screen "D_Bar_1" 1280x800
   Bar "Static" at 6,4 size 40x120
   TextField "Label_Static" at 6,156 size 55x22; Text 'Static'
   Bar "A_Range" at 98,4 size 40x120
      Appearance <- "D_Range"
   TextField "Label_A_Range" at 98,156 size 79x22; Text 'A_Range'
   Bar "A_Flash" at 190,4 size 40x120
      Appearance <- "D_Range"
   TextField "Label_A_Flash" at 190,156 size 72x22; Text 'A_Flash'
   Bar "A_Bit" at 282,4 size 40x120
      Appearance <- "D_Bool"
   TextField "Label_A_Bit" at 282,156 size 51x22; Text 'A_Bit'
   Bar "A_Bits" at 374,4 size 40x120
      Appearance <- "D_Bits"
   TextField "Label_A_Bits" at 374,156 size 60x22; Text 'A_Bits'
   Bar "V_Range" at 466,4 size 40x120
      Visibility <- "D_Range"
   TextField "Label_V_Range" at 466,156 size 79x22; Text 'V_Range'
   Bar "V_Bit" at 558,4 size 40x120
      Visibility <- "D_Vis"
   TextField "Label_V_Bit" at 558,156 size 51x22; Text 'V_Bit'
   Bar "M_H" at 650,4 size 40x120
      HorizontalMovement <- "D_Pct"
   TextField "Label_M_H" at 650,156 size 42x22; Text 'M_H'
   Bar "M_V" at 742,4 size 40x120
      VerticalMovement <- "D_Pct"
   TextField "Label_M_V" at 742,156 size 41x22; Text 'M_V'
   Bar "M_D" at 834,4 size 40x120
      DiagonalMovement <- "D_Pct"
   TextField "Label_M_D" at 834,156 size 42x22; Text 'M_D'
   Bar "M_Direct" at 926,4 size 40x120
      DirectMovement <- "D_X"
      DirectMovement <- "D_Y"
   TextField "Label_M_Direct" at 926,156 size 82x22; Text 'M_Direct'
   Bar "E_Range" at 1018,4 size 40x120
      ObjectEnable <- "D_Range"
   TextField "Label_E_Range" at 1018,156 size 78x22; Text 'E_Range'
   Bar "E_Bit" at 1110,4 size 40x120
      ObjectEnable <- "D_En"
   TextField "Label_E_Bit" at 1110,156 size 50x22; Text 'E_Bit'
   Bar "PV_Pct" at 6,176 size 40x120
      ProcessValue <- "D_Pct"
   TextField "Label_PV_Pct" at 6,328 size 65x22; Text 'PV_Pct'
   Bar "PV_Real" at 98,176 size 40x120
      ProcessValue <- "D_Real"
   TextField "Label_PV_Real" at 98,328 size 76x22; Text 'PV_Real'
   Bar "PV_BarR" at 190,176 size 40x120
      ProcessValue <- "D_BarR"
   TextField "Label_PV_BarR" at 190,328 size 79x22; Text 'PV_BarR'
   Bar "PV_Pct_0_100" at 282,176 size 40x120; MinimumValue 0; MaximumValue 100
      ProcessValue <- "D_Pct"
   TextField "Label_PV_Pct_0_100" at 282,328 size 131x22; Text 'PV_Pct_0_100'
   Bar "PV_Pct_MaxMin" at 374,176 size 40x120
      ProcessValue <- "D_Pct"
      MaximumValue <- "D_Max"
      MinimumValue <- "D_Min"
   TextField "Label_PV_Pct_MaxMin" at 374,328 size 140x22; Text 'PV_Pct_MaxMin'
   IOField "State" at 4,774 size 60x22; FormatPattern 9
      ProcessValue <- "D_State"
   Button "S1" at 70,774 size 40x22; TextOff 'S1'
      on Click: "SetS1"()
   Button "S2" at 114,774 size 40x22; TextOff 'S2'
      on Click: "SetS2"()
   Button "S3" at 158,774 size 40x22; TextOff 'S3'
      on Click: "SetS3"()
   Button "S4" at 202,774 size 40x22; TextOff 'S4'
      on Click: "SetS4"()
   Button "Next" at 1236,774 size 40x22; TextOff 'Next'
      on Click: ActivateScreen("D_Switch_1", 0)

screen "D_Button_1" 1280x800
   Button "Static" at 6,4 size 100x40; TextOff 'Text'
   TextField "Label_Static" at 6,76 size 55x22; Text 'Static'
   Button "A_Range" at 158,4 size 100x40; TextOff 'Text'
      Appearance <- "D_Range"
   TextField "Label_A_Range" at 158,76 size 79x22; Text 'A_Range'
   Button "A_Flash" at 310,4 size 100x40; TextOff 'Text'
      Appearance <- "D_Range"
   TextField "Label_A_Flash" at 310,76 size 72x22; Text 'A_Flash'
   Button "A_Bit" at 462,4 size 100x40; TextOff 'Text'
      Appearance <- "D_Bool"
   TextField "Label_A_Bit" at 462,76 size 51x22; Text 'A_Bit'
   Button "A_Bits" at 614,4 size 100x40; TextOff 'Text'
      Appearance <- "D_Bits"
   TextField "Label_A_Bits" at 614,76 size 60x22; Text 'A_Bits'
   Button "V_Range" at 766,4 size 100x40; TextOff 'Text'
      Visibility <- "D_Range"
   TextField "Label_V_Range" at 766,76 size 79x22; Text 'V_Range'
   Button "V_Bit" at 918,4 size 100x40; TextOff 'Text'
      Visibility <- "D_Vis"
   TextField "Label_V_Bit" at 918,76 size 51x22; Text 'V_Bit'
   Button "M_H" at 1070,4 size 100x40; TextOff 'Text'
      HorizontalMovement <- "D_Pct"
   TextField "Label_M_H" at 1070,76 size 42x22; Text 'M_H'
   Button "M_V" at 6,96 size 100x40; TextOff 'Text'
      VerticalMovement <- "D_Pct"
   TextField "Label_M_V" at 6,168 size 41x22; Text 'M_V'
   Button "M_D" at 158,96 size 100x40; TextOff 'Text'
      DiagonalMovement <- "D_Pct"
   TextField "Label_M_D" at 158,168 size 42x22; Text 'M_D'
   Button "M_Direct" at 310,96 size 100x40; TextOff 'Text'
      DirectMovement <- "D_X"
      DirectMovement <- "D_Y"
   TextField "Label_M_Direct" at 310,168 size 82x22; Text 'M_Direct'
   Button "E_Range" at 462,96 size 100x40; TextOff 'Text'
      ObjectEnable <- "D_Range"
   TextField "Label_E_Range" at 462,168 size 78x22; Text 'E_Range'
   Button "E_Bit" at 614,96 size 100x40; TextOff 'Text'
      ObjectEnable <- "D_En"
   TextField "Label_E_Bit" at 614,168 size 50x22; Text 'E_Bit'
   IOField "State" at 4,774 size 60x22; FormatPattern 9
      ProcessValue <- "D_State"
   Button "S1" at 70,774 size 40x22; TextOff 'S1'
      on Click: "SetS1"()
   Button "S2" at 114,774 size 40x22; TextOff 'S2'
      on Click: "SetS2"()
   Button "S3" at 158,774 size 40x22; TextOff 'S3'
      on Click: "SetS3"()
   Button "S4" at 202,774 size 40x22; TextOff 'S4'
      on Click: "SetS4"()
   Button "Next" at 1236,774 size 40x22; TextOff 'Next'
      on Click: ActivateScreen("D_SymbolicIOField_1", 0)

screen "D_Circle_1" 1280x800
   TextField "Label_Static" at 6,86 size 55x22; Text 'Static'
   Circle "A_Range" at 108,4 size 50x50
      Appearance <- "D_Range"
   TextField "Label_A_Range" at 108,86 size 79x22; Text 'A_Range'
   Circle "A_Flash" at 210,4 size 50x50
      Appearance <- "D_Range"
   TextField "Label_A_Flash" at 210,86 size 72x22; Text 'A_Flash'
   Circle "A_Bit" at 312,4 size 50x50
      Appearance <- "D_Bool"
   TextField "Label_A_Bit" at 312,86 size 51x22; Text 'A_Bit'
   Circle "A_Bits" at 414,4 size 50x50
      Appearance <- "D_Bits"
   TextField "Label_A_Bits" at 414,86 size 60x22; Text 'A_Bits'
   Circle "V_Range" at 516,4 size 50x50
      Visibility <- "D_Range"
   TextField "Label_V_Range" at 516,86 size 79x22; Text 'V_Range'
   Circle "V_Bit" at 618,4 size 50x50
      Visibility <- "D_Vis"
   TextField "Label_V_Bit" at 618,86 size 51x22; Text 'V_Bit'
   Circle "M_H" at 720,4 size 50x50
      HorizontalMovement <- "D_Pct"
   TextField "Label_M_H" at 720,86 size 42x22; Text 'M_H'
   Circle "M_V" at 822,4 size 50x50
      VerticalMovement <- "D_Pct"
   TextField "Label_M_V" at 822,86 size 41x22; Text 'M_V'
   Circle "M_D" at 924,4 size 50x50
      DiagonalMovement <- "D_Pct"
   TextField "Label_M_D" at 924,86 size 42x22; Text 'M_D'
   Circle "M_Direct" at 1026,4 size 50x50
      DirectMovement <- "D_X"
      DirectMovement <- "D_Y"
   TextField "Label_M_Direct" at 1026,86 size 82x22; Text 'M_Direct'
   Circle "E_Range" at 1128,4 size 50x50
      ObjectEnable <- "D_Range"
   TextField "Label_E_Range" at 1128,86 size 78x22; Text 'E_Range'
   Circle "E_Bit" at 6,106 size 50x50
      ObjectEnable <- "D_En"
   TextField "Label_E_Bit" at 6,188 size 50x22; Text 'E_Bit'
   IOField "State" at 4,774 size 60x22; FormatPattern 9
      ProcessValue <- "D_State"
   Button "S1" at 70,774 size 40x22; TextOff 'S1'
      on Click: "SetS1"()
   Button "S2" at 114,774 size 40x22; TextOff 'S2'
      on Click: "SetS2"()
   Button "S3" at 158,774 size 40x22; TextOff 'S3'
      on Click: "SetS3"()
   Button "S4" at 202,774 size 40x22; TextOff 'S4'
      on Click: "SetS4"()
   Button "Next" at 1236,774 size 40x22; TextOff 'Next'
      on Click: ActivateScreen("D_Rectangle_1", 0)

screen "D_Clock_1" 1280x800
   Clock "Static" at 6,4 size 150x150
   TextField "Label_Static" at 6,186 size 55x22; Text 'Static'
   Clock "A_Range" at 208,4 size 150x150
      Appearance <- "D_Range"
   TextField "Label_A_Range" at 208,186 size 79x22; Text 'A_Range'
   Clock "A_Flash" at 410,4 size 150x150
      Appearance <- "D_Range"
   TextField "Label_A_Flash" at 410,186 size 72x22; Text 'A_Flash'
   Clock "A_Bit" at 612,4 size 150x150
      Appearance <- "D_Bool"
   TextField "Label_A_Bit" at 612,186 size 51x22; Text 'A_Bit'
   Clock "A_Bits" at 814,4 size 150x150
      Appearance <- "D_Bits"
   TextField "Label_A_Bits" at 814,186 size 60x22; Text 'A_Bits'
   Clock "V_Range" at 1016,4 size 150x150
      Visibility <- "D_Range"
   TextField "Label_V_Range" at 1016,186 size 79x22; Text 'V_Range'
   Clock "V_Bit" at 6,206 size 150x150
      Visibility <- "D_Vis"
   TextField "Label_V_Bit" at 6,388 size 51x22; Text 'V_Bit'
   Clock "M_H" at 208,206 size 150x150
      HorizontalMovement <- "D_Pct"
   TextField "Label_M_H" at 208,388 size 42x22; Text 'M_H'
   Clock "M_V" at 410,206 size 150x150
      VerticalMovement <- "D_Pct"
   TextField "Label_M_V" at 410,388 size 41x22; Text 'M_V'
   Clock "M_D" at 612,206 size 150x150
      DiagonalMovement <- "D_Pct"
   TextField "Label_M_D" at 612,388 size 42x22; Text 'M_D'
   Clock "M_Direct" at 814,206 size 150x150
      DirectMovement <- "D_X"
      DirectMovement <- "D_Y"
   TextField "Label_M_Direct" at 814,388 size 82x22; Text 'M_Direct'
   Clock "E_Range" at 1016,206 size 150x150
      ObjectEnable <- "D_Range"
   TextField "Label_E_Range" at 1016,388 size 78x22; Text 'E_Range'
   Clock "E_Bit" at 6,408 size 150x150
      ObjectEnable <- "D_En"
   TextField "Label_E_Bit" at 6,590 size 50x22; Text 'E_Bit'
   IOField "State" at 4,774 size 60x22; FormatPattern 9
      ProcessValue <- "D_State"
   Button "S1" at 70,774 size 40x22; TextOff 'S1'
      on Click: "SetS1"()
   Button "S2" at 114,774 size 40x22; TextOff 'S2'
      on Click: "SetS2"()
   Button "S3" at 158,774 size 40x22; TextOff 'S3'
      on Click: "SetS3"()
   Button "S4" at 202,774 size 40x22; TextOff 'S4'
      on Click: "SetS4"()
   Button "Next" at 1236,774 size 40x22; TextOff 'Next'
      on Click: ActivateScreen("D_Line_1", 0)

screen "D_DateTimeField_1" 1280x800
   DateTimeField "Static" at 6,4 size 189x26
   TextField "Label_Static" at 6,66 size 55x22; Text 'Static'
   DateTimeField "A_Range" at 218,4 size 189x26
      Appearance <- "D_Range"
   TextField "Label_A_Range" at 218,66 size 79x22; Text 'A_Range'
   DateTimeField "A_Flash" at 430,4 size 189x26
      Appearance <- "D_Range"
   TextField "Label_A_Flash" at 430,66 size 72x22; Text 'A_Flash'
   DateTimeField "A_Bit" at 642,4 size 189x26
      Appearance <- "D_Bool"
   TextField "Label_A_Bit" at 642,66 size 51x22; Text 'A_Bit'
   DateTimeField "A_Bits" at 854,4 size 189x26
      Appearance <- "D_Bits"
   TextField "Label_A_Bits" at 854,66 size 60x22; Text 'A_Bits'
   DateTimeField "V_Range" at 1066,4 size 189x26
      Visibility <- "D_Range"
   TextField "Label_V_Range" at 1066,66 size 79x22; Text 'V_Range'
   DateTimeField "V_Bit" at 6,86 size 189x26
      Visibility <- "D_Vis"
   TextField "Label_V_Bit" at 6,148 size 51x22; Text 'V_Bit'
   DateTimeField "M_H" at 218,86 size 189x26
      HorizontalMovement <- "D_Pct"
   TextField "Label_M_H" at 218,148 size 42x22; Text 'M_H'
   DateTimeField "M_V" at 430,86 size 189x26
      VerticalMovement <- "D_Pct"
   TextField "Label_M_V" at 430,148 size 41x22; Text 'M_V'
   DateTimeField "M_D" at 642,86 size 189x26
      DiagonalMovement <- "D_Pct"
   TextField "Label_M_D" at 642,148 size 42x22; Text 'M_D'
   DateTimeField "M_Direct" at 854,86 size 189x26
      DirectMovement <- "D_X"
      DirectMovement <- "D_Y"
   TextField "Label_M_Direct" at 854,148 size 82x22; Text 'M_Direct'
   DateTimeField "E_Range" at 1066,86 size 189x26
      ObjectEnable <- "D_Range"
   TextField "Label_E_Range" at 1066,148 size 78x22; Text 'E_Range'
   DateTimeField "E_Bit" at 6,168 size 189x26
      ObjectEnable <- "D_En"
   TextField "Label_E_Bit" at 6,230 size 50x22; Text 'E_Bit'
   DateTimeField "PV_DateTime" at 218,168 size 189x26
      ProcessValue <- "D_DateTime"
   TextField "Label_PV_DateTime" at 218,230 size 117x22; Text 'PV_DateTime'
   IOField "State" at 4,774 size 60x22; FormatPattern 9
      ProcessValue <- "D_State"
   Button "S1" at 70,774 size 40x22; TextOff 'S1'
      on Click: "SetS1"()
   Button "S2" at 114,774 size 40x22; TextOff 'S2'
      on Click: "SetS2"()
   Button "S3" at 158,774 size 40x22; TextOff 'S3'
      on Click: "SetS3"()
   Button "S4" at 202,774 size 40x22; TextOff 'S4'
      on Click: "SetS4"()
   Button "Next" at 1236,774 size 40x22; TextOff 'Next'
      on Click: ActivateScreen("D_Bar_1", 0)

screen "D_Ellipse_1" 1280x800
   TextField "Label_Static" at 6,86 size 55x22; Text 'Static'
   Ellipse "A_Range" at 158,4 size 100x50
      Appearance <- "D_Range"
   TextField "Label_A_Range" at 158,86 size 79x22; Text 'A_Range'
   Ellipse "A_Flash" at 310,4 size 100x50
      Appearance <- "D_Range"
   TextField "Label_A_Flash" at 310,86 size 72x22; Text 'A_Flash'
   Ellipse "A_Bit" at 462,4 size 100x50
      Appearance <- "D_Bool"
   TextField "Label_A_Bit" at 462,86 size 51x22; Text 'A_Bit'
   Ellipse "A_Bits" at 614,4 size 100x50
      Appearance <- "D_Bits"
   TextField "Label_A_Bits" at 614,86 size 60x22; Text 'A_Bits'
   Ellipse "V_Range" at 766,4 size 100x50
      Visibility <- "D_Range"
   TextField "Label_V_Range" at 766,86 size 79x22; Text 'V_Range'
   Ellipse "V_Bit" at 918,4 size 100x50
      Visibility <- "D_Vis"
   TextField "Label_V_Bit" at 918,86 size 51x22; Text 'V_Bit'
   Ellipse "M_H" at 1070,4 size 100x50
      HorizontalMovement <- "D_Pct"
   TextField "Label_M_H" at 1070,86 size 42x22; Text 'M_H'
   Ellipse "M_V" at 6,106 size 100x50
      VerticalMovement <- "D_Pct"
   TextField "Label_M_V" at 6,188 size 41x22; Text 'M_V'
   Ellipse "M_D" at 158,106 size 100x50
      DiagonalMovement <- "D_Pct"
   TextField "Label_M_D" at 158,188 size 42x22; Text 'M_D'
   Ellipse "M_Direct" at 310,106 size 100x50
      DirectMovement <- "D_X"
      DirectMovement <- "D_Y"
   TextField "Label_M_Direct" at 310,188 size 82x22; Text 'M_Direct'
   Ellipse "E_Range" at 462,106 size 100x50
      ObjectEnable <- "D_Range"
   TextField "Label_E_Range" at 462,188 size 78x22; Text 'E_Range'
   Ellipse "E_Bit" at 614,106 size 100x50
      ObjectEnable <- "D_En"
   TextField "Label_E_Bit" at 614,188 size 50x22; Text 'E_Bit'
   IOField "State" at 4,774 size 60x22; FormatPattern 9
      ProcessValue <- "D_State"
   Button "S1" at 70,774 size 40x22; TextOff 'S1'
      on Click: "SetS1"()
   Button "S2" at 114,774 size 40x22; TextOff 'S2'
      on Click: "SetS2"()
   Button "S3" at 158,774 size 40x22; TextOff 'S3'
      on Click: "SetS3"()
   Button "S4" at 202,774 size 40x22; TextOff 'S4'
      on Click: "SetS4"()
   Button "Next" at 1236,774 size 40x22; TextOff 'Next'
      on Click: ActivateScreen("D_Circle_1", 0)

screen "D_Gauge_1" 1280x800
   Gauge "Static" at 6,4 size 150x150; CaptionText 'SIMATIC'
   TextField "Label_Static" at 6,186 size 55x22; Text 'Static'
   Gauge "A_Range" at 208,4 size 150x150; CaptionText 'SIMATIC'
      Appearance <- "D_Range"
   TextField "Label_A_Range" at 208,186 size 79x22; Text 'A_Range'
   Gauge "A_Flash" at 410,4 size 150x150; CaptionText 'SIMATIC'
      Appearance <- "D_Range"
   TextField "Label_A_Flash" at 410,186 size 72x22; Text 'A_Flash'
   Gauge "A_Bit" at 612,4 size 150x150; CaptionText 'SIMATIC'
      Appearance <- "D_Bool"
   TextField "Label_A_Bit" at 612,186 size 51x22; Text 'A_Bit'
   Gauge "A_Bits" at 814,4 size 150x150; CaptionText 'SIMATIC'
      Appearance <- "D_Bits"
   TextField "Label_A_Bits" at 814,186 size 60x22; Text 'A_Bits'
   Gauge "V_Range" at 1016,4 size 150x150; CaptionText 'SIMATIC'
      Visibility <- "D_Range"
   TextField "Label_V_Range" at 1016,186 size 79x22; Text 'V_Range'
   Gauge "V_Bit" at 6,206 size 150x150; CaptionText 'SIMATIC'
      Visibility <- "D_Vis"
   TextField "Label_V_Bit" at 6,388 size 51x22; Text 'V_Bit'
   Gauge "M_H" at 208,206 size 150x150; CaptionText 'SIMATIC'
      HorizontalMovement <- "D_Pct"
   TextField "Label_M_H" at 208,388 size 42x22; Text 'M_H'
   Gauge "M_V" at 410,206 size 150x150; CaptionText 'SIMATIC'
      VerticalMovement <- "D_Pct"
   TextField "Label_M_V" at 410,388 size 41x22; Text 'M_V'
   Gauge "M_D" at 612,206 size 150x150; CaptionText 'SIMATIC'
      DiagonalMovement <- "D_Pct"
   TextField "Label_M_D" at 612,388 size 42x22; Text 'M_D'
   Gauge "M_Direct" at 814,206 size 150x150; CaptionText 'SIMATIC'
      DirectMovement <- "D_X"
      DirectMovement <- "D_Y"
   TextField "Label_M_Direct" at 814,388 size 82x22; Text 'M_Direct'
   Gauge "E_Range" at 1016,206 size 150x150; CaptionText 'SIMATIC'
      ObjectEnable <- "D_Range"
   TextField "Label_E_Range" at 1016,388 size 78x22; Text 'E_Range'
   Gauge "E_Bit" at 6,408 size 150x150; CaptionText 'SIMATIC'
      ObjectEnable <- "D_En"
   TextField "Label_E_Bit" at 6,590 size 50x22; Text 'E_Bit'
   Gauge "PV_Pct" at 208,408 size 150x150; CaptionText 'SIMATIC'
      ProcessValue <- "D_Pct"
   TextField "Label_PV_Pct" at 208,590 size 65x22; Text 'PV_Pct'
   Gauge "PV_Real" at 410,408 size 150x150; CaptionText 'SIMATIC'
      ProcessValue <- "D_Real"
   TextField "Label_PV_Real" at 410,590 size 76x22; Text 'PV_Real'
   Gauge "PV_Pct_MaxMin" at 612,408 size 150x150; CaptionText 'SIMATIC'
      ProcessValue <- "D_Pct"
      MaximumValue <- "D_Max"
      MinimumValue <- "D_Min"
   TextField "Label_PV_Pct_MaxMin" at 612,590 size 140x22; Text 'PV_Pct_MaxMin'
   IOField "State" at 4,774 size 60x22; FormatPattern 9
      ProcessValue <- "D_State"
   Button "S1" at 70,774 size 40x22; TextOff 'S1'
      on Click: "SetS1"()
   Button "S2" at 114,774 size 40x22; TextOff 'S2'
      on Click: "SetS2"()
   Button "S3" at 158,774 size 40x22; TextOff 'S3'
      on Click: "SetS3"()
   Button "S4" at 202,774 size 40x22; TextOff 'S4'
      on Click: "SetS4"()
   Button "Next" at 1236,774 size 40x22; TextOff 'Next'
      on Click: ActivateScreen("D_Clock_1", 0)

screen "D_GraphicIOField_1" 1280x800
   GraphicIOField "Static" at 6,4 size 60x60
   TextField "Label_Static" at 6,96 size 55x22; Text 'Static'
   GraphicIOField "A_Range" at 118,4 size 60x60
      Appearance <- "D_Range"
   TextField "Label_A_Range" at 118,96 size 79x22; Text 'A_Range'
   GraphicIOField "A_Flash" at 230,4 size 60x60
      Appearance <- "D_Range"
   TextField "Label_A_Flash" at 230,96 size 72x22; Text 'A_Flash'
   GraphicIOField "A_Bit" at 342,4 size 60x60
      Appearance <- "D_Bool"
   TextField "Label_A_Bit" at 342,96 size 51x22; Text 'A_Bit'
   GraphicIOField "A_Bits" at 454,4 size 60x60
      Appearance <- "D_Bits"
   TextField "Label_A_Bits" at 454,96 size 60x22; Text 'A_Bits'
   GraphicIOField "V_Range" at 566,4 size 60x60
      Visibility <- "D_Range"
   TextField "Label_V_Range" at 566,96 size 79x22; Text 'V_Range'
   GraphicIOField "V_Bit" at 678,4 size 60x60
      Visibility <- "D_Vis"
   TextField "Label_V_Bit" at 678,96 size 51x22; Text 'V_Bit'
   GraphicIOField "M_H" at 790,4 size 60x60
      HorizontalMovement <- "D_Pct"
   TextField "Label_M_H" at 790,96 size 42x22; Text 'M_H'
   GraphicIOField "M_V" at 902,4 size 60x60
      VerticalMovement <- "D_Pct"
   TextField "Label_M_V" at 902,96 size 41x22; Text 'M_V'
   GraphicIOField "M_D" at 1014,4 size 60x60
      DiagonalMovement <- "D_Pct"
   TextField "Label_M_D" at 1014,96 size 42x22; Text 'M_D'
   GraphicIOField "M_Direct" at 1126,4 size 60x60
      DirectMovement <- "D_X"
      DirectMovement <- "D_Y"
   TextField "Label_M_Direct" at 1126,96 size 82x22; Text 'M_Direct'
   GraphicIOField "E_Range" at 6,116 size 60x60
      ObjectEnable <- "D_Range"
   TextField "Label_E_Range" at 6,208 size 78x22; Text 'E_Range'
   GraphicIOField "E_Bit" at 118,116 size 60x60
      ObjectEnable <- "D_En"
   TextField "Label_E_Bit" at 118,208 size 50x22; Text 'E_Bit'
   IOField "State" at 4,774 size 60x22; FormatPattern 9
      ProcessValue <- "D_State"
   Button "S1" at 70,774 size 40x22; TextOff 'S1'
      on Click: "SetS1"()
   Button "S2" at 114,774 size 40x22; TextOff 'S2'
      on Click: "SetS2"()
   Button "S3" at 158,774 size 40x22; TextOff 'S3'
      on Click: "SetS3"()
   Button "S4" at 202,774 size 40x22; TextOff 'S4'
      on Click: "SetS4"()
   Button "Next" at 1236,774 size 40x22; TextOff 'Next'
      on Click: ActivateScreen("D_DateTimeField_1", 0)

screen "D_GraphicView_1" 1280x800
   GraphicView "Static" at 6,4 size 100x60
   TextField "Label_Static" at 6,96 size 55x22; Text 'Static'
   GraphicView "A_Range" at 158,4 size 100x60
      Appearance <- "D_Range"
   TextField "Label_A_Range" at 158,96 size 79x22; Text 'A_Range'
   GraphicView "A_Flash" at 310,4 size 100x60
      Appearance <- "D_Range"
   TextField "Label_A_Flash" at 310,96 size 72x22; Text 'A_Flash'
   GraphicView "A_Bit" at 462,4 size 100x60
      Appearance <- "D_Bool"
   TextField "Label_A_Bit" at 462,96 size 51x22; Text 'A_Bit'
   GraphicView "A_Bits" at 614,4 size 100x60
      Appearance <- "D_Bits"
   TextField "Label_A_Bits" at 614,96 size 60x22; Text 'A_Bits'
   GraphicView "V_Range" at 766,4 size 100x60
      Visibility <- "D_Range"
   TextField "Label_V_Range" at 766,96 size 79x22; Text 'V_Range'
   GraphicView "V_Bit" at 918,4 size 100x60
      Visibility <- "D_Vis"
   TextField "Label_V_Bit" at 918,96 size 51x22; Text 'V_Bit'
   GraphicView "M_H" at 1070,4 size 100x60
      HorizontalMovement <- "D_Pct"
   TextField "Label_M_H" at 1070,96 size 42x22; Text 'M_H'
   GraphicView "M_V" at 6,116 size 100x60
      VerticalMovement <- "D_Pct"
   TextField "Label_M_V" at 6,208 size 41x22; Text 'M_V'
   GraphicView "M_D" at 158,116 size 100x60
      DiagonalMovement <- "D_Pct"
   TextField "Label_M_D" at 158,208 size 42x22; Text 'M_D'
   GraphicView "M_Direct" at 310,116 size 100x60
      DirectMovement <- "D_X"
      DirectMovement <- "D_Y"
   TextField "Label_M_Direct" at 310,208 size 82x22; Text 'M_Direct'
   GraphicView "E_Range" at 462,116 size 100x60
      ObjectEnable <- "D_Range"
   TextField "Label_E_Range" at 462,208 size 78x22; Text 'E_Range'
   GraphicView "E_Bit" at 614,116 size 100x60
      ObjectEnable <- "D_En"
   TextField "Label_E_Bit" at 614,208 size 50x22; Text 'E_Bit'
   IOField "State" at 4,774 size 60x22; FormatPattern 9
      ProcessValue <- "D_State"
   Button "S1" at 70,774 size 40x22; TextOff 'S1'
      on Click: "SetS1"()
   Button "S2" at 114,774 size 40x22; TextOff 'S2'
      on Click: "SetS2"()
   Button "S3" at 158,774 size 40x22; TextOff 'S3'
      on Click: "SetS3"()
   Button "S4" at 202,774 size 40x22; TextOff 'S4'
      on Click: "SetS4"()
   Button "Next" at 1236,774 size 40x22; TextOff 'Next'
      on Click: ActivateScreen("D_IOField_1", 0)

screen "D_IOField_1" 1280x800
   IOField "Static" at 6,4 size 100x30
   TextField "Label_Static" at 6,66 size 55x22; Text 'Static'
   IOField "A_Range" at 158,4 size 100x30
      Appearance <- "D_Range"
   TextField "Label_A_Range" at 158,66 size 79x22; Text 'A_Range'
   IOField "A_Flash" at 310,4 size 100x30
      Appearance <- "D_Range"
   TextField "Label_A_Flash" at 310,66 size 72x22; Text 'A_Flash'
   IOField "A_Bit" at 462,4 size 100x30
      Appearance <- "D_Bool"
   TextField "Label_A_Bit" at 462,66 size 51x22; Text 'A_Bit'
   IOField "A_Bits" at 614,4 size 100x30
      Appearance <- "D_Bits"
   TextField "Label_A_Bits" at 614,66 size 60x22; Text 'A_Bits'
   IOField "V_Range" at 766,4 size 100x30
      Visibility <- "D_Range"
   TextField "Label_V_Range" at 766,66 size 79x22; Text 'V_Range'
   IOField "V_Bit" at 918,4 size 100x30
      Visibility <- "D_Vis"
   TextField "Label_V_Bit" at 918,66 size 51x22; Text 'V_Bit'
   IOField "M_H" at 1070,4 size 100x30
      HorizontalMovement <- "D_Pct"
   TextField "Label_M_H" at 1070,66 size 42x22; Text 'M_H'
   IOField "M_V" at 6,86 size 100x30
      VerticalMovement <- "D_Pct"
   TextField "Label_M_V" at 6,148 size 41x22; Text 'M_V'
   IOField "M_D" at 158,86 size 100x30
      DiagonalMovement <- "D_Pct"
   TextField "Label_M_D" at 158,148 size 42x22; Text 'M_D'
   IOField "M_Direct" at 310,86 size 100x30
      DirectMovement <- "D_X"
      DirectMovement <- "D_Y"
   TextField "Label_M_Direct" at 310,148 size 82x22; Text 'M_Direct'
   IOField "E_Range" at 462,86 size 100x30
      ObjectEnable <- "D_Range"
   TextField "Label_E_Range" at 462,148 size 78x22; Text 'E_Range'
   IOField "E_Bit" at 614,86 size 100x30
      ObjectEnable <- "D_En"
   TextField "Label_E_Bit" at 614,148 size 50x22; Text 'E_Bit'
   IOField "PV_SInt" at 766,86 size 100x30; FormatPattern s999
      ProcessValue <- "D_SInt"
   TextField "Label_PV_SInt" at 766,148 size 74x22; Text 'PV_SInt'
   IOField "PV_Int" at 918,86 size 100x30; FormatPattern s99999
      ProcessValue <- "D_Int"
   TextField "Label_PV_Int" at 918,148 size 63x22; Text 'PV_Int'
   IOField "PV_DInt" at 1070,86 size 100x30; FormatPattern s9999999999
      ProcessValue <- "D_DInt"
   TextField "Label_PV_DInt" at 1070,148 size 75x22; Text 'PV_DInt'
   IOField "PV_USInt" at 6,168 size 100x30; FormatPattern 999
      ProcessValue <- "D_USInt"
   TextField "Label_PV_USInt" at 6,230 size 86x22; Text 'PV_USInt'
   IOField "PV_UInt" at 158,168 size 100x30; FormatPattern 99999
      ProcessValue <- "D_UInt"
   TextField "Label_PV_UInt" at 158,230 size 75x22; Text 'PV_UInt'
   IOField "PV_UDInt" at 310,168 size 100x30; FormatPattern 9999999999
      ProcessValue <- "D_UDInt"
   TextField "Label_PV_UDInt" at 310,230 size 87x22; Text 'PV_UDInt'
   IOField "PV_Real" at 462,168 size 100x30
      ProcessValue <- "D_Real"
   TextField "Label_PV_Real" at 462,230 size 76x22; Text 'PV_Real'
   IOField "PV_LReal" at 614,168 size 100x30
      ProcessValue <- "D_LReal"
   TextField "Label_PV_LReal" at 614,230 size 86x22; Text 'PV_LReal'
   IOField "PV_String" at 766,168 size 100x30
      ProcessValue <- "D_String"
   TextField "Label_PV_String" at 766,230 size 90x22; Text 'PV_String'
   IOField "PV_Int_Shift2" at 918,168 size 100x30; FormatPattern s99999
      ProcessValue <- "D_Int"
   TextField "Label_PV_Int_Shift2" at 918,230 size 126x22; Text 'PV_Int_Shift2'
   IOField "PV_Int_s999999" at 1070,168 size 100x30; FormatPattern s999999
      ProcessValue <- "D_Int"
   TextField "Label_PV_Int_s999999" at 1070,230 size 149x22; Text 'PV_Int_s999999'
   IOField "PV_Real_s9999_99" at 6,250 size 100x30; FormatPattern s9999.99
      ProcessValue <- "D_Real"
   TextField "Label_PV_Real_s9999_99" at 6,312 size 173x22; Text 'PV_Real_s9999_99'
   IOField "PV_Int_Output" at 158,250 size 100x30; FormatPattern s99999
      ProcessValue <- "D_Int"
   TextField "Label_PV_Int_Output" at 158,312 size 131x22; Text 'PV_Int_Output'
   IOField "PV_Int_s99" at 310,250 size 100x30; FormatPattern s99
      ProcessValue <- "D_Int"
   TextField "Label_PV_Int_s99" at 310,312 size 105x22; Text 'PV_Int_s99'
   IOField "State" at 4,774 size 60x22; FormatPattern 9
      ProcessValue <- "D_State"
   Button "S1" at 70,774 size 40x22; TextOff 'S1'
      on Click: "SetS1"()
   Button "S2" at 114,774 size 40x22; TextOff 'S2'
      on Click: "SetS2"()
   Button "S3" at 158,774 size 40x22; TextOff 'S3'
      on Click: "SetS3"()
   Button "S4" at 202,774 size 40x22; TextOff 'S4'
      on Click: "SetS4"()
   Button "Next" at 1236,774 size 40x22; TextOff 'Next'
      on Click: ActivateScreen("D_Button_1", 0)

screen "D_Line_1" 1280x800
   TextField "Label_Static" at 6,86 size 55x22; Text 'Static'
   Line "A_Range" at 158,4 size 100x50
      Appearance <- "D_Range"
   TextField "Label_A_Range" at 158,86 size 79x22; Text 'A_Range'
   Line "A_Flash" at 310,4 size 100x50
      Appearance <- "D_Range"
   TextField "Label_A_Flash" at 310,86 size 72x22; Text 'A_Flash'
   Line "A_Bit" at 462,4 size 100x50
      Appearance <- "D_Bool"
   TextField "Label_A_Bit" at 462,86 size 51x22; Text 'A_Bit'
   Line "A_Bits" at 614,4 size 100x50
      Appearance <- "D_Bits"
   TextField "Label_A_Bits" at 614,86 size 60x22; Text 'A_Bits'
   Line "V_Range" at 766,4 size 100x50
      Visibility <- "D_Range"
   TextField "Label_V_Range" at 766,86 size 79x22; Text 'V_Range'
   Line "V_Bit" at 918,4 size 100x50
      Visibility <- "D_Vis"
   TextField "Label_V_Bit" at 918,86 size 51x22; Text 'V_Bit'
   Line "M_H" at 1070,4 size 100x50
      HorizontalMovement <- "D_Pct"
   TextField "Label_M_H" at 1070,86 size 42x22; Text 'M_H'
   Line "M_V" at 6,106 size 100x50
      VerticalMovement <- "D_Pct"
   TextField "Label_M_V" at 6,188 size 41x22; Text 'M_V'
   Line "M_D" at 158,106 size 100x50
      DiagonalMovement <- "D_Pct"
   TextField "Label_M_D" at 158,188 size 42x22; Text 'M_D'
   Line "M_Direct" at 310,106 size 100x50
      DirectMovement <- "D_X"
      DirectMovement <- "D_Y"
   TextField "Label_M_Direct" at 310,188 size 82x22; Text 'M_Direct'
   Line "E_Range" at 462,106 size 100x50
      ObjectEnable <- "D_Range"
   TextField "Label_E_Range" at 462,188 size 78x22; Text 'E_Range'
   Line "E_Bit" at 614,106 size 100x50
      ObjectEnable <- "D_En"
   TextField "Label_E_Bit" at 614,188 size 50x22; Text 'E_Bit'
   IOField "State" at 4,774 size 60x22; FormatPattern 9
      ProcessValue <- "D_State"
   Button "S1" at 70,774 size 40x22; TextOff 'S1'
      on Click: "SetS1"()
   Button "S2" at 114,774 size 40x22; TextOff 'S2'
      on Click: "SetS2"()
   Button "S3" at 158,774 size 40x22; TextOff 'S3'
      on Click: "SetS3"()
   Button "S4" at 202,774 size 40x22; TextOff 'S4'
      on Click: "SetS4"()
   Button "Next" at 1236,774 size 40x22; TextOff 'Next'
      on Click: ActivateScreen("D_Polyline_1", 0)

screen "D_Polygon_1" 1280x800
   TextField "Label_Static" at 6,86 size 55x22; Text 'Static'
   Polygon "A_Range" at 158,4 size 100x50
      Appearance <- "D_Range"
   TextField "Label_A_Range" at 158,86 size 79x22; Text 'A_Range'
   Polygon "A_Flash" at 310,4 size 100x50
      Appearance <- "D_Range"
   TextField "Label_A_Flash" at 310,86 size 72x22; Text 'A_Flash'
   Polygon "A_Bit" at 462,4 size 100x50
      Appearance <- "D_Bool"
   TextField "Label_A_Bit" at 462,86 size 51x22; Text 'A_Bit'
   Polygon "A_Bits" at 614,4 size 100x50
      Appearance <- "D_Bits"
   TextField "Label_A_Bits" at 614,86 size 60x22; Text 'A_Bits'
   Polygon "V_Range" at 766,4 size 100x50
      Visibility <- "D_Range"
   TextField "Label_V_Range" at 766,86 size 79x22; Text 'V_Range'
   Polygon "V_Bit" at 918,4 size 100x50
      Visibility <- "D_Vis"
   TextField "Label_V_Bit" at 918,86 size 51x22; Text 'V_Bit'
   Polygon "M_H" at 1070,4 size 100x50
      HorizontalMovement <- "D_Pct"
   TextField "Label_M_H" at 1070,86 size 42x22; Text 'M_H'
   Polygon "M_V" at 6,106 size 100x50
      VerticalMovement <- "D_Pct"
   TextField "Label_M_V" at 6,188 size 41x22; Text 'M_V'
   Polygon "M_D" at 158,106 size 100x50
      DiagonalMovement <- "D_Pct"
   TextField "Label_M_D" at 158,188 size 42x22; Text 'M_D'
   Polygon "M_Direct" at 310,106 size 100x50
      DirectMovement <- "D_X"
      DirectMovement <- "D_Y"
   TextField "Label_M_Direct" at 310,188 size 82x22; Text 'M_Direct'
   Polygon "E_Range" at 462,106 size 100x50
      ObjectEnable <- "D_Range"
   TextField "Label_E_Range" at 462,188 size 78x22; Text 'E_Range'
   Polygon "E_Bit" at 614,106 size 100x50
      ObjectEnable <- "D_En"
   TextField "Label_E_Bit" at 614,188 size 50x22; Text 'E_Bit'
   IOField "State" at 4,774 size 60x22; FormatPattern 9
      ProcessValue <- "D_State"
   Button "S1" at 70,774 size 40x22; TextOff 'S1'
      on Click: "SetS1"()
   Button "S2" at 114,774 size 40x22; TextOff 'S2'
      on Click: "SetS2"()
   Button "S3" at 158,774 size 40x22; TextOff 'S3'
      on Click: "SetS3"()
   Button "S4" at 202,774 size 40x22; TextOff 'S4'
      on Click: "SetS4"()
   Button "Next" at 1236,774 size 40x22; TextOff 'Next'
      on Click: ActivateScreen("D_Ellipse_1", 0)

screen "D_Polyline_1" 1280x800
   TextField "Label_Static" at 6,86 size 55x22; Text 'Static'
   Polyline "A_Range" at 158,4 size 100x50
      Appearance <- "D_Range"
   TextField "Label_A_Range" at 158,86 size 79x22; Text 'A_Range'
   Polyline "A_Flash" at 310,4 size 100x50
      Appearance <- "D_Range"
   TextField "Label_A_Flash" at 310,86 size 72x22; Text 'A_Flash'
   Polyline "A_Bit" at 462,4 size 100x50
      Appearance <- "D_Bool"
   TextField "Label_A_Bit" at 462,86 size 51x22; Text 'A_Bit'
   Polyline "A_Bits" at 614,4 size 100x50
      Appearance <- "D_Bits"
   TextField "Label_A_Bits" at 614,86 size 60x22; Text 'A_Bits'
   Polyline "V_Range" at 766,4 size 100x50
      Visibility <- "D_Range"
   TextField "Label_V_Range" at 766,86 size 79x22; Text 'V_Range'
   Polyline "V_Bit" at 918,4 size 100x50
      Visibility <- "D_Vis"
   TextField "Label_V_Bit" at 918,86 size 51x22; Text 'V_Bit'
   Polyline "M_H" at 1070,4 size 100x50
      HorizontalMovement <- "D_Pct"
   TextField "Label_M_H" at 1070,86 size 42x22; Text 'M_H'
   Polyline "M_V" at 6,106 size 100x50
      VerticalMovement <- "D_Pct"
   TextField "Label_M_V" at 6,188 size 41x22; Text 'M_V'
   Polyline "M_D" at 158,106 size 100x50
      DiagonalMovement <- "D_Pct"
   TextField "Label_M_D" at 158,188 size 42x22; Text 'M_D'
   Polyline "M_Direct" at 310,106 size 100x50
      DirectMovement <- "D_X"
      DirectMovement <- "D_Y"
   TextField "Label_M_Direct" at 310,188 size 82x22; Text 'M_Direct'
   Polyline "E_Range" at 462,106 size 100x50
      ObjectEnable <- "D_Range"
   TextField "Label_E_Range" at 462,188 size 78x22; Text 'E_Range'
   Polyline "E_Bit" at 614,106 size 100x50
      ObjectEnable <- "D_En"
   TextField "Label_E_Bit" at 614,188 size 50x22; Text 'E_Bit'
   IOField "State" at 4,774 size 60x22; FormatPattern 9
      ProcessValue <- "D_State"
   Button "S1" at 70,774 size 40x22; TextOff 'S1'
      on Click: "SetS1"()
   Button "S2" at 114,774 size 40x22; TextOff 'S2'
      on Click: "SetS2"()
   Button "S3" at 158,774 size 40x22; TextOff 'S3'
      on Click: "SetS3"()
   Button "S4" at 202,774 size 40x22; TextOff 'S4'
      on Click: "SetS4"()
   Button "Next" at 1236,774 size 40x22; TextOff 'Next'
      on Click: ActivateScreen("D_Polygon_1", 0)

screen "D_Rectangle_1" 1280x800
   TextField "Label_Static" at 6,86 size 55x22; Text 'Static'
   Rectangle "A_Range" at 158,4 size 100x50
      Appearance <- "D_Range"
   TextField "Label_A_Range" at 158,86 size 79x22; Text 'A_Range'
   Rectangle "A_Flash" at 310,4 size 100x50
      Appearance <- "D_Range"
   TextField "Label_A_Flash" at 310,86 size 72x22; Text 'A_Flash'
   Rectangle "A_Bit" at 462,4 size 100x50
      Appearance <- "D_Bool"
   TextField "Label_A_Bit" at 462,86 size 51x22; Text 'A_Bit'
   Rectangle "A_Bits" at 614,4 size 100x50
      Appearance <- "D_Bits"
   TextField "Label_A_Bits" at 614,86 size 60x22; Text 'A_Bits'
   Rectangle "V_Range" at 766,4 size 100x50
      Visibility <- "D_Range"
   TextField "Label_V_Range" at 766,86 size 79x22; Text 'V_Range'
   Rectangle "V_Bit" at 918,4 size 100x50
      Visibility <- "D_Vis"
   TextField "Label_V_Bit" at 918,86 size 51x22; Text 'V_Bit'
   Rectangle "M_H" at 1070,4 size 100x50
      HorizontalMovement <- "D_Pct"
   TextField "Label_M_H" at 1070,86 size 42x22; Text 'M_H'
   Rectangle "M_V" at 6,106 size 100x50
      VerticalMovement <- "D_Pct"
   TextField "Label_M_V" at 6,188 size 41x22; Text 'M_V'
   Rectangle "M_D" at 158,106 size 100x50
      DiagonalMovement <- "D_Pct"
   TextField "Label_M_D" at 158,188 size 42x22; Text 'M_D'
   Rectangle "M_Direct" at 310,106 size 100x50
      DirectMovement <- "D_X"
      DirectMovement <- "D_Y"
   TextField "Label_M_Direct" at 310,188 size 82x22; Text 'M_Direct'
   Rectangle "E_Range" at 462,106 size 100x50
      ObjectEnable <- "D_Range"
   TextField "Label_E_Range" at 462,188 size 78x22; Text 'E_Range'
   Rectangle "E_Bit" at 614,106 size 100x50
      ObjectEnable <- "D_En"
   TextField "Label_E_Bit" at 614,188 size 50x22; Text 'E_Bit'
   IOField "State" at 4,774 size 60x22; FormatPattern 9
      ProcessValue <- "D_State"
   Button "S1" at 70,774 size 40x22; TextOff 'S1'
      on Click: "SetS1"()
   Button "S2" at 114,774 size 40x22; TextOff 'S2'
      on Click: "SetS2"()
   Button "S3" at 158,774 size 40x22; TextOff 'S3'
      on Click: "SetS3"()
   Button "S4" at 202,774 size 40x22; TextOff 'S4'
      on Click: "SetS4"()
   Button "Next" at 1236,774 size 40x22; TextOff 'Next'
      on Click: ActivateScreen("D_TextField_1", 0)

screen "D_Slider_1" 1280x800
   Slider "Static" at 6,4 size 60x160; Caption 'SIMATIC'
   TextField "Label_Static" at 6,196 size 55x22; Text 'Static'
   Slider "A_Range" at 118,4 size 60x160; Caption 'SIMATIC'
      Appearance <- "D_Range"
   TextField "Label_A_Range" at 118,196 size 79x22; Text 'A_Range'
   Slider "A_Flash" at 230,4 size 60x160; Caption 'SIMATIC'
      Appearance <- "D_Range"
   TextField "Label_A_Flash" at 230,196 size 72x22; Text 'A_Flash'
   Slider "A_Bit" at 342,4 size 60x160; Caption 'SIMATIC'
      Appearance <- "D_Bool"
   TextField "Label_A_Bit" at 342,196 size 51x22; Text 'A_Bit'
   Slider "A_Bits" at 454,4 size 60x160; Caption 'SIMATIC'
      Appearance <- "D_Bits"
   TextField "Label_A_Bits" at 454,196 size 60x22; Text 'A_Bits'
   Slider "V_Range" at 566,4 size 60x160; Caption 'SIMATIC'
      Visibility <- "D_Range"
   TextField "Label_V_Range" at 566,196 size 79x22; Text 'V_Range'
   Slider "V_Bit" at 678,4 size 60x160; Caption 'SIMATIC'
      Visibility <- "D_Vis"
   TextField "Label_V_Bit" at 678,196 size 51x22; Text 'V_Bit'
   Slider "M_H" at 790,4 size 60x160; Caption 'SIMATIC'
      HorizontalMovement <- "D_Pct"
   TextField "Label_M_H" at 790,196 size 42x22; Text 'M_H'
   Slider "M_V" at 902,4 size 60x160; Caption 'SIMATIC'
      VerticalMovement <- "D_Pct"
   TextField "Label_M_V" at 902,196 size 41x22; Text 'M_V'
   Slider "M_D" at 1014,4 size 60x160; Caption 'SIMATIC'
      DiagonalMovement <- "D_Pct"
   TextField "Label_M_D" at 1014,196 size 42x22; Text 'M_D'
   Slider "M_Direct" at 1126,4 size 60x160; Caption 'SIMATIC'
      DirectMovement <- "D_X"
      DirectMovement <- "D_Y"
   TextField "Label_M_Direct" at 1126,196 size 82x22; Text 'M_Direct'
   Slider "E_Range" at 6,216 size 60x160; Caption 'SIMATIC'
      ObjectEnable <- "D_Range"
   TextField "Label_E_Range" at 6,408 size 78x22; Text 'E_Range'
   Slider "E_Bit" at 118,216 size 60x160; Caption 'SIMATIC'
      ObjectEnable <- "D_En"
   TextField "Label_E_Bit" at 118,408 size 50x22; Text 'E_Bit'
   Slider "PV_Pct" at 230,216 size 60x160; Caption 'SIMATIC'
      ProcessValue <- "D_Pct"
   TextField "Label_PV_Pct" at 230,408 size 65x22; Text 'PV_Pct'
   Slider "PV_Int" at 342,216 size 60x160; Caption 'SIMATIC'
      ProcessValue <- "D_Int"
   TextField "Label_PV_Int" at 342,408 size 63x22; Text 'PV_Int'
   Slider "PV_Pct_0_200" at 454,216 size 60x160; Caption 'SIMATIC'
      ProcessValue <- "D_Pct"
   TextField "Label_PV_Pct_0_200" at 454,408 size 131x22; Text 'PV_Pct_0_200'
   IOField "State" at 4,774 size 60x22; FormatPattern 9
      ProcessValue <- "D_State"
   Button "S1" at 70,774 size 40x22; TextOff 'S1'
      on Click: "SetS1"()
   Button "S2" at 114,774 size 40x22; TextOff 'S2'
      on Click: "SetS2"()
   Button "S3" at 158,774 size 40x22; TextOff 'S3'
      on Click: "SetS3"()
   Button "S4" at 202,774 size 40x22; TextOff 'S4'
      on Click: "SetS4"()
   Button "Next" at 1236,774 size 40x22; TextOff 'Next'
      on Click: ActivateScreen("D_Gauge_1", 0)

screen "D_Switch_1" 1280x800
   Switch "Static" at 6,4 size 120x40; CaptionText 'Switch'; TextOff '0'; TextOn '1'
   TextField "Label_Static" at 6,76 size 55x22; Text 'Static'
   Switch "A_Range" at 178,4 size 120x40; CaptionText 'Switch'; TextOff '0'; TextOn '1'
      Appearance <- "D_Range"
   TextField "Label_A_Range" at 178,76 size 79x22; Text 'A_Range'
   Switch "A_Flash" at 350,4 size 120x40; CaptionText 'Switch'; TextOff '0'; TextOn '1'
      Appearance <- "D_Range"
   TextField "Label_A_Flash" at 350,76 size 72x22; Text 'A_Flash'
   Switch "A_Bit" at 522,4 size 120x40; CaptionText 'Switch'; TextOff '0'; TextOn '1'
      Appearance <- "D_Bool"
   TextField "Label_A_Bit" at 522,76 size 51x22; Text 'A_Bit'
   Switch "A_Bits" at 694,4 size 120x40; CaptionText 'Switch'; TextOff '0'; TextOn '1'
      Appearance <- "D_Bits"
   TextField "Label_A_Bits" at 694,76 size 60x22; Text 'A_Bits'
   Switch "V_Range" at 866,4 size 120x40; CaptionText 'Switch'; TextOff '0'; TextOn '1'
      Visibility <- "D_Range"
   TextField "Label_V_Range" at 866,76 size 79x22; Text 'V_Range'
   Switch "V_Bit" at 1038,4 size 120x40; CaptionText 'Switch'; TextOff '0'; TextOn '1'
      Visibility <- "D_Vis"
   TextField "Label_V_Bit" at 1038,76 size 51x22; Text 'V_Bit'
   Switch "M_H" at 6,96 size 120x40; CaptionText 'Switch'; TextOff '0'; TextOn '1'
      HorizontalMovement <- "D_Pct"
   TextField "Label_M_H" at 6,168 size 42x22; Text 'M_H'
   Switch "M_V" at 178,96 size 120x40; CaptionText 'Switch'; TextOff '0'; TextOn '1'
      VerticalMovement <- "D_Pct"
   TextField "Label_M_V" at 178,168 size 41x22; Text 'M_V'
   Switch "M_D" at 350,96 size 120x40; CaptionText 'Switch'; TextOff '0'; TextOn '1'
      DiagonalMovement <- "D_Pct"
   TextField "Label_M_D" at 350,168 size 42x22; Text 'M_D'
   Switch "M_Direct" at 522,96 size 120x40; CaptionText 'Switch'; TextOff '0'; TextOn '1'
      DirectMovement <- "D_X"
      DirectMovement <- "D_Y"
   TextField "Label_M_Direct" at 522,168 size 82x22; Text 'M_Direct'
   Switch "E_Range" at 694,96 size 120x40; CaptionText 'Switch'; TextOff '0'; TextOn '1'
      ObjectEnable <- "D_Range"
   TextField "Label_E_Range" at 694,168 size 78x22; Text 'E_Range'
   Switch "E_Bit" at 866,96 size 120x40; CaptionText 'Switch'; TextOff '0'; TextOn '1'
      ObjectEnable <- "D_En"
   TextField "Label_E_Bit" at 866,168 size 50x22; Text 'E_Bit'
   Switch "PV_Bool" at 1038,96 size 120x40; CaptionText 'Switch'; TextOff '0'; TextOn '1'
      ProcessValue <- "D_Bool"
   TextField "Label_PV_Bool" at 1038,168 size 75x22; Text 'PV_Bool'
   IOField "State" at 4,774 size 60x22; FormatPattern 9
      ProcessValue <- "D_State"
   Button "S1" at 70,774 size 40x22; TextOff 'S1'
      on Click: "SetS1"()
   Button "S2" at 114,774 size 40x22; TextOff 'S2'
      on Click: "SetS2"()
   Button "S3" at 158,774 size 40x22; TextOff 'S3'
      on Click: "SetS3"()
   Button "S4" at 202,774 size 40x22; TextOff 'S4'
      on Click: "SetS4"()
   Button "Next" at 1236,774 size 40x22; TextOff 'Next'
      on Click: ActivateScreen("D_SymbolLibrary_1", 0)

screen "D_SymbolicIOField_1" 1280x800
   SymbolicIOField "Static" at 6,4 size 120x30; TextOff '0'; TextOn '1'
   TextField "Label_Static" at 6,66 size 55x22; Text 'Static'
   SymbolicIOField "A_Range" at 178,4 size 120x30; TextOff '0'; TextOn '1'
      Appearance <- "D_Range"
   TextField "Label_A_Range" at 178,66 size 79x22; Text 'A_Range'
   SymbolicIOField "A_Flash" at 350,4 size 120x30; TextOff '0'; TextOn '1'
      Appearance <- "D_Range"
   TextField "Label_A_Flash" at 350,66 size 72x22; Text 'A_Flash'
   SymbolicIOField "A_Bit" at 522,4 size 120x30; TextOff '0'; TextOn '1'
      Appearance <- "D_Bool"
   TextField "Label_A_Bit" at 522,66 size 51x22; Text 'A_Bit'
   SymbolicIOField "A_Bits" at 694,4 size 120x30; TextOff '0'; TextOn '1'
      Appearance <- "D_Bits"
   TextField "Label_A_Bits" at 694,66 size 60x22; Text 'A_Bits'
   SymbolicIOField "V_Range" at 866,4 size 120x30; TextOff '0'; TextOn '1'
      Visibility <- "D_Range"
   TextField "Label_V_Range" at 866,66 size 79x22; Text 'V_Range'
   SymbolicIOField "V_Bit" at 1038,4 size 120x30; TextOff '0'; TextOn '1'
      Visibility <- "D_Vis"
   TextField "Label_V_Bit" at 1038,66 size 51x22; Text 'V_Bit'
   SymbolicIOField "M_H" at 6,86 size 120x30; TextOff '0'; TextOn '1'
      HorizontalMovement <- "D_Pct"
   TextField "Label_M_H" at 6,148 size 42x22; Text 'M_H'
   SymbolicIOField "M_V" at 178,86 size 120x30; TextOff '0'; TextOn '1'
      VerticalMovement <- "D_Pct"
   TextField "Label_M_V" at 178,148 size 41x22; Text 'M_V'
   SymbolicIOField "M_D" at 350,86 size 120x30; TextOff '0'; TextOn '1'
      DiagonalMovement <- "D_Pct"
   TextField "Label_M_D" at 350,148 size 42x22; Text 'M_D'
   SymbolicIOField "M_Direct" at 522,86 size 120x30; TextOff '0'; TextOn '1'
      DirectMovement <- "D_X"
      DirectMovement <- "D_Y"
   TextField "Label_M_Direct" at 522,148 size 82x22; Text 'M_Direct'
   SymbolicIOField "E_Range" at 694,86 size 120x30; TextOff '0'; TextOn '1'
      ObjectEnable <- "D_Range"
   TextField "Label_E_Range" at 694,148 size 78x22; Text 'E_Range'
   SymbolicIOField "E_Bit" at 866,86 size 120x30; TextOff '0'; TextOn '1'
      ObjectEnable <- "D_En"
   TextField "Label_E_Bit" at 866,148 size 50x22; Text 'E_Bit'
   SymbolicIOField "PV_TL_Value" at 1038,86 size 120x30; TextOff '0'; TextOn '1'; TextList "TL_Value"
      ProcessValue <- "D_TL"
   TextField "Label_PV_TL_Value" at 1038,148 size 116x22; Text 'PV_TL_Value'
   SymbolicIOField "PV_TL_Bit" at 6,168 size 120x30; TextOff '0'; TextOn '1'; TextList "TL_Bit"
      ProcessValue <- "D_Bool"
   TextField "Label_PV_TL_Bit" at 6,230 size 93x22; Text 'PV_TL_Bit'
   SymbolicIOField "PV_TL_BitNo" at 178,168 size 120x30; TextOff '0'; TextOn '1'; TextList "TL_BitNo"
      ProcessValue <- "D_Bits"
   TextField "Label_PV_TL_BitNo" at 178,230 size 116x22; Text 'PV_TL_BitNo'
   IOField "State" at 4,774 size 60x22; FormatPattern 9
      ProcessValue <- "D_State"
   Button "S1" at 70,774 size 40x22; TextOff 'S1'
      on Click: "SetS1"()
   Button "S2" at 114,774 size 40x22; TextOff 'S2'
      on Click: "SetS2"()
   Button "S3" at 158,774 size 40x22; TextOff 'S3'
      on Click: "SetS3"()
   Button "S4" at 202,774 size 40x22; TextOff 'S4'
      on Click: "SetS4"()
   Button "Next" at 1236,774 size 40x22; TextOff 'Next'
      on Click: ActivateScreen("D_GraphicIOField_1", 0)

screen "D_SymbolLibrary_1" 1280x800
   SymbolLibrary "Static" at 6,4 size 60x60
   TextField "Label_Static" at 6,96 size 55x22; Text 'Static'
   SymbolLibrary "A_Range" at 118,4 size 60x60
      Appearance <- "D_Range"
   TextField "Label_A_Range" at 118,96 size 79x22; Text 'A_Range'
   SymbolLibrary "A_Flash" at 230,4 size 60x60
      Appearance <- "D_Range"
   TextField "Label_A_Flash" at 230,96 size 72x22; Text 'A_Flash'
   SymbolLibrary "A_Bit" at 342,4 size 60x60
      Appearance <- "D_Bool"
   TextField "Label_A_Bit" at 342,96 size 51x22; Text 'A_Bit'
   SymbolLibrary "A_Bits" at 454,4 size 60x60
      Appearance <- "D_Bits"
   TextField "Label_A_Bits" at 454,96 size 60x22; Text 'A_Bits'
   SymbolLibrary "V_Range" at 566,4 size 60x60
      Visibility <- "D_Range"
   TextField "Label_V_Range" at 566,96 size 79x22; Text 'V_Range'
   SymbolLibrary "V_Bit" at 678,4 size 60x60
      Visibility <- "D_Vis"
   TextField "Label_V_Bit" at 678,96 size 51x22; Text 'V_Bit'
   SymbolLibrary "M_H" at 790,4 size 60x60
      HorizontalMovement <- "D_Pct"
   TextField "Label_M_H" at 790,96 size 42x22; Text 'M_H'
   SymbolLibrary "M_V" at 902,4 size 60x60
      VerticalMovement <- "D_Pct"
   TextField "Label_M_V" at 902,96 size 41x22; Text 'M_V'
   SymbolLibrary "M_D" at 1014,4 size 60x60
      DiagonalMovement <- "D_Pct"
   TextField "Label_M_D" at 1014,96 size 42x22; Text 'M_D'
   SymbolLibrary "M_Direct" at 1126,4 size 60x60
      DirectMovement <- "D_X"
      DirectMovement <- "D_Y"
   TextField "Label_M_Direct" at 1126,96 size 82x22; Text 'M_Direct'
   SymbolLibrary "E_Range" at 6,116 size 60x60
      ObjectEnable <- "D_Range"
   TextField "Label_E_Range" at 6,208 size 78x22; Text 'E_Range'
   SymbolLibrary "E_Bit" at 118,116 size 60x60
      ObjectEnable <- "D_En"
   TextField "Label_E_Bit" at 118,208 size 50x22; Text 'E_Bit'
   SymbolLibrary "PV_Pct" at 230,116 size 60x60
      ProcessValue <- "D_Pct"
   TextField "Label_PV_Pct" at 230,208 size 65x22; Text 'PV_Pct'
   IOField "State" at 4,774 size 60x22; FormatPattern 9
      ProcessValue <- "D_State"
   Button "S1" at 70,774 size 40x22; TextOff 'S1'
      on Click: "SetS1"()
   Button "S2" at 114,774 size 40x22; TextOff 'S2'
      on Click: "SetS2"()
   Button "S3" at 158,774 size 40x22; TextOff 'S3'
      on Click: "SetS3"()
   Button "S4" at 202,774 size 40x22; TextOff 'S4'
      on Click: "SetS4"()
   Button "Next" at 1236,774 size 40x22; TextOff 'Next'
      on Click: ActivateScreen("D_Slider_1", 0)

screen "D_TextField_1" 1280x800
   TextField "Static" at 6,4 size 42x22; Text 'Text'
   TextField "Label_Static" at 6,66 size 55x22; Text 'Static'
   TextField "A_Range" at 158,4 size 42x22; Text 'Text'
      Appearance <- "D_Range"
   TextField "Label_A_Range" at 158,66 size 79x22; Text 'A_Range'
   TextField "A_Flash" at 310,4 size 42x22; Text 'Text'
      Appearance <- "D_Range"
   TextField "Label_A_Flash" at 310,66 size 72x22; Text 'A_Flash'
   TextField "A_Bit" at 462,4 size 42x22; Text 'Text'
      Appearance <- "D_Bool"
   TextField "Label_A_Bit" at 462,66 size 51x22; Text 'A_Bit'
   TextField "A_Bits" at 614,4 size 42x22; Text 'Text'
      Appearance <- "D_Bits"
   TextField "Label_A_Bits" at 614,66 size 60x22; Text 'A_Bits'
   TextField "V_Range" at 766,4 size 42x22; Text 'Text'
      Visibility <- "D_Range"
   TextField "Label_V_Range" at 766,66 size 79x22; Text 'V_Range'
   TextField "V_Bit" at 918,4 size 42x22; Text 'Text'
      Visibility <- "D_Vis"
   TextField "Label_V_Bit" at 918,66 size 51x22; Text 'V_Bit'
   TextField "M_H" at 1070,4 size 42x22; Text 'Text'
      HorizontalMovement <- "D_Pct"
   TextField "Label_M_H" at 1070,66 size 42x22; Text 'M_H'
   TextField "M_V" at 6,86 size 42x22; Text 'Text'
      VerticalMovement <- "D_Pct"
   TextField "Label_M_V" at 6,148 size 41x22; Text 'M_V'
   TextField "M_D" at 158,86 size 42x22; Text 'Text'
      DiagonalMovement <- "D_Pct"
   TextField "Label_M_D" at 158,148 size 42x22; Text 'M_D'
   TextField "M_Direct" at 310,86 size 42x22; Text 'Text'
      DirectMovement <- "D_X"
      DirectMovement <- "D_Y"
   TextField "Label_M_Direct" at 310,148 size 82x22; Text 'M_Direct'
   TextField "E_Range" at 462,86 size 42x22; Text 'Text'
      ObjectEnable <- "D_Range"
   TextField "Label_E_Range" at 462,148 size 78x22; Text 'E_Range'
   TextField "E_Bit" at 614,86 size 42x22; Text 'Text'
      ObjectEnable <- "D_En"
   TextField "Label_E_Bit" at 614,148 size 50x22; Text 'E_Bit'
   IOField "State" at 4,774 size 60x22; FormatPattern 9
      ProcessValue <- "D_State"
   Button "S1" at 70,774 size 40x22; TextOff 'S1'
      on Click: "SetS1"()
   Button "S2" at 114,774 size 40x22; TextOff 'S2'
      on Click: "SetS2"()
   Button "S3" at 158,774 size 40x22; TextOff 'S3'
      on Click: "SetS3"()
   Button "S4" at 202,774 size 40x22; TextOff 'S4'
      on Click: "SetS4"()
   Button "Next" at 1236,774 size 40x22; TextOff 'Next'
      on Click: ActivateScreen("D_GraphicView_1", 0)

screen "C5_Buttons" 1280x800, template "T_C05"
   Button "Btn_Text" at 6,40 size 120x50; TextOff 'Btn_Text off'; TextOn 'Btn_Text on'
   TextField "Label_Btn_Text" at 6,92 size 81x22; Text 'Btn_Text'
   Button "Btn_Graphic" at 182,40 size 120x90; TextOff 'Btn_Graphic off'; TextOn 'Btn_Graphic on'; PictureOff "G_PNG"; PictureOn "G_JPG"
   TextField "Label_Btn_Graphic" at 182,132 size 109x22; Text 'Btn_Graphic'
   Button "Btn_GraphicAndText" at 358,40 size 120x90; TextOff 'Btn_GraphicAndText off'; TextOn 'Btn_GraphicAndText on'; PictureOff "G_SVG"; PictureOn "G_EMF"
   TextField "Label_Btn_GraphicAndText" at 358,132 size 177x22; Text 'Btn_GraphicAndText'
   Button "Btn_TextList" at 534,40 size 160x50; TextOff 'Btn_TextList off'; TextOn 'Btn_TextList on'; TextList "TL_Value"
      ProcessValue <- "D_TL"
   TextField "Label_Btn_TextList" at 534,92 size 113x22; Text 'Btn_TextList'
   Button "Btn_GraphicList" at 710,40 size 120x90; TextOff 'Btn_GraphicList off'; TextOn 'Btn_GraphicList on'; PictureList "GL_Value"
      ProcessValue <- "D_TL"
   TextField "Label_Btn_GraphicList" at 710,132 size 141x22; Text 'Btn_GraphicList'
   Button "Btn_Invisible" at 886,40 size 120x50; TextOff 'Btn_Invisible off'; TextOn 'Btn_Invisible on'
   TextField "Label_Btn_Invisible" at 886,92 size 119x22; Text 'Btn_Invisible'
   Switch "Sw_Switch" at 1062,40 size 120x40; CaptionText 'Switch'; TextOff '0'; TextOn '1'
      ProcessValue <- "D_Bool"
   TextField "Label_Sw_Switch" at 1062,82 size 98x22; Text 'Sw_Switch'
   Switch "Sw_Text" at 6,152 size 120x40; CaptionText 'Switch'; TextOff 'Sw_Text off'; TextOn 'Sw_Text on'
      ProcessValue <- "D_Bool"
   TextField "Label_Sw_Text" at 6,194 size 78x22; Text 'Sw_Text'
   Switch "Sw_Graphic" at 182,152 size 120x90; CaptionText 'Switch'; TextOff '0'; TextOn '1'; PictureOff "G_BMP"; PictureOn "G_GIF"
      ProcessValue <- "D_Bool"
   TextField "Label_Sw_Graphic" at 182,244 size 106x22; Text 'Sw_Graphic'
   IOField "State" at 4,774 size 60x22; FormatPattern 9
      ProcessValue <- "D_State"
   Button "S1" at 70,774 size 40x22; TextOff 'S1'
      on Click: "SetS1"()
   Button "S2" at 114,774 size 40x22; TextOff 'S2'
      on Click: "SetS2"()
   Button "S3" at 158,774 size 40x22; TextOff 'S3'
      on Click: "SetS3"()
   Button "S4" at 202,774 size 40x22; TextOff 'S4'
      on Click: "SetS4"()
   Button "Next" at 1236,774 size 40x22; TextOff 'Next'
      on Click: ActivateScreen("C5_Structure", 0)

screen "C5_GraphicView_1" 1280x800, template "T_C05"
   GraphicView "GV_PNG" at 6,40 size 120x80; Picture "G_PNG"
   TextField "Label_GV_PNG" at 6,122 size 75x22; Text 'GV_PNG'
   GraphicView "GV_JPG" at 142,40 size 120x80; Picture "G_JPG"
   TextField "Label_GV_JPG" at 142,122 size 71x22; Text 'GV_JPG'
   GraphicView "GV_BMP" at 278,40 size 120x80; Picture "G_BMP"
   TextField "Label_GV_BMP" at 278,122 size 75x22; Text 'GV_BMP'
   GraphicView "GV_GIF" at 414,40 size 120x80; Picture "G_GIF"
   TextField "Label_GV_GIF" at 414,122 size 69x22; Text 'GV_GIF'
   GraphicView "GV_TIF" at 550,40 size 120x80; Picture "G_TIF"
   TextField "Label_GV_TIF" at 550,122 size 67x22; Text 'GV_TIF'
   GraphicView "GV_EMF" at 686,40 size 120x80; Picture "G_EMF"
   TextField "Label_GV_EMF" at 686,122 size 73x22; Text 'GV_EMF'
   GraphicView "GV_WMF" at 822,40 size 120x80; Picture "G_WMF"
   TextField "Label_GV_WMF" at 822,122 size 79x22; Text 'GV_WMF'
   GraphicView "GV_SVG" at 958,40 size 120x80; Picture "G_SVG"
   TextField "Label_GV_SVG" at 958,122 size 73x22; Text 'GV_SVG'
   GraphicView "GV_TALL" at 1094,40 size 120x80; Picture "G_TALL"
   TextField "Label_GV_TALL" at 1094,122 size 80x22; Text 'GV_TALL'
   GraphicView "GV_WIDE" at 6,142 size 120x80; Picture "G_WIDE"
   TextField "Label_GV_WIDE" at 6,224 size 85x22; Text 'GV_WIDE'
   IOField "State" at 4,774 size 60x22; FormatPattern 9
      ProcessValue <- "D_State"
   Button "S1" at 70,774 size 40x22; TextOff 'S1'
      on Click: "SetS1"()
   Button "S2" at 114,774 size 40x22; TextOff 'S2'
      on Click: "SetS2"()
   Button "S3" at 158,774 size 40x22; TextOff 'S3'
      on Click: "SetS3"()
   Button "S4" at 202,774 size 40x22; TextOff 'S4'
      on Click: "SetS4"()
   Button "Next" at 1236,774 size 40x22; TextOff 'Next'
      on Click: ActivateScreen("C5_GraphicView_2", 0)

screen "C5_GraphicView_2" 1280x800, template "T_C05"
   GraphicView "PNG_160x60_FitF" at 6,40 size 160x60; Picture "G_PNG"
   TextField "Label_PNG_160x60_FitF" at 6,102 size 161x22; Text 'PNG_160x60_FitF'
   GraphicView "PNG_160x60_FitT" at 182,40 size 160x60; Picture "G_PNG"
   TextField "Label_PNG_160x60_FitT" at 182,102 size 161x22; Text 'PNG_160x60_FitT'
   GraphicView "PNG_60x120_FitF" at 358,40 size 60x120; Picture "G_PNG"
   TextField "Label_PNG_60x120_FitF" at 358,162 size 161x22; Text 'PNG_60x120_FitF'
   GraphicView "PNG_60x120_FitT" at 534,40 size 60x120; Picture "G_PNG"
   TextField "Label_PNG_60x120_FitT" at 534,162 size 161x22; Text 'PNG_60x120_FitT'
   GraphicView "PNG_80x80_FitF" at 710,40 size 80x80; Picture "G_PNG"
   TextField "Label_PNG_80x80_FitF" at 710,122 size 150x22; Text 'PNG_80x80_FitF'
   GraphicView "PNG_80x80_FitT" at 886,40 size 80x80; Picture "G_PNG"
   TextField "Label_PNG_80x80_FitT" at 886,122 size 150x22; Text 'PNG_80x80_FitT'
   GraphicView "TALL_160x60_FitF" at 1062,40 size 160x60; Picture "G_TALL"
   TextField "Label_TALL_160x60_FitF" at 1062,102 size 166x22; Text 'TALL_160x60_FitF'
   GraphicView "TALL_160x60_FitT" at 6,182 size 160x60; Picture "G_TALL"
   TextField "Label_TALL_160x60_FitT" at 6,244 size 166x22; Text 'TALL_160x60_FitT'
   GraphicView "TALL_60x120_FitF" at 182,182 size 60x120; Picture "G_TALL"
   TextField "Label_TALL_60x120_FitF" at 182,304 size 166x22; Text 'TALL_60x120_FitF'
   GraphicView "TALL_60x120_FitT" at 358,182 size 60x120; Picture "G_TALL"
   TextField "Label_TALL_60x120_FitT" at 358,304 size 166x22; Text 'TALL_60x120_FitT'
   GraphicView "TALL_80x80_FitF" at 534,182 size 80x80; Picture "G_TALL"
   TextField "Label_TALL_80x80_FitF" at 534,264 size 155x22; Text 'TALL_80x80_FitF'
   GraphicView "TALL_80x80_FitT" at 710,182 size 80x80; Picture "G_TALL"
   TextField "Label_TALL_80x80_FitT" at 710,264 size 155x22; Text 'TALL_80x80_FitT'
   GraphicView "WIDE_160x60_FitF" at 886,182 size 160x60; Picture "G_WIDE"
   TextField "Label_WIDE_160x60_FitF" at 886,244 size 171x22; Text 'WIDE_160x60_FitF'
   GraphicView "WIDE_160x60_FitT" at 1062,182 size 160x60; Picture "G_WIDE"
   TextField "Label_WIDE_160x60_FitT" at 1062,244 size 171x22; Text 'WIDE_160x60_FitT'
   GraphicView "WIDE_60x120_FitF" at 6,324 size 60x120; Picture "G_WIDE"
   TextField "Label_WIDE_60x120_FitF" at 6,446 size 171x22; Text 'WIDE_60x120_FitF'
   GraphicView "WIDE_60x120_FitT" at 182,324 size 60x120; Picture "G_WIDE"
   TextField "Label_WIDE_60x120_FitT" at 182,446 size 171x22; Text 'WIDE_60x120_FitT'
   GraphicView "WIDE_80x80_FitF" at 358,324 size 80x80; Picture "G_WIDE"
   TextField "Label_WIDE_80x80_FitF" at 358,406 size 160x22; Text 'WIDE_80x80_FitF'
   GraphicView "WIDE_80x80_FitT" at 534,324 size 80x80; Picture "G_WIDE"
   TextField "Label_WIDE_80x80_FitT" at 534,406 size 160x22; Text 'WIDE_80x80_FitT'
   GraphicView "BMP_Transparent" at 710,324 size 120x80; Picture "G_BMP"
   TextField "Label_BMP_Transparent" at 710,406 size 154x22; Text 'BMP_Transparent'
   GraphicView "PNG_BackTransparent" at 886,324 size 120x80; Picture "G_PNG"
   TextField "Label_PNG_BackTransparent" at 886,406 size 194x22; Text 'PNG_BackTransparent'
   IOField "State" at 4,774 size 60x22; FormatPattern 9
      ProcessValue <- "D_State"
   Button "S1" at 70,774 size 40x22; TextOff 'S1'
      on Click: "SetS1"()
   Button "S2" at 114,774 size 40x22; TextOff 'S2'
      on Click: "SetS2"()
   Button "S3" at 158,774 size 40x22; TextOff 'S3'
      on Click: "SetS3"()
   Button "S4" at 202,774 size 40x22; TextOff 'S4'
      on Click: "SetS4"()
   Button "Next" at 1236,774 size 40x22; TextOff 'Next'
      on Click: ActivateScreen("C5_Lists", 0)

screen "C5_Lists" 1280x800, template "T_C05"
   SymbolicIOField "SIO_TL_Value" at 6,40 size 160x30; TextOff '0'; TextOn '1'; TextList "TL_Value"
      ProcessValue <- "D_TL"
   TextField "Label_SIO_TL_Value" at 6,72 size 126x22; Text 'SIO_TL_Value'
   SymbolicIOField "SIO_TL_Bit" at 182,40 size 160x30; TextOff '0'; TextOn '1'; TextList "TL_Bit"
      ProcessValue <- "D_Bool"
   TextField "Label_SIO_TL_Bit" at 182,72 size 103x22; Text 'SIO_TL_Bit'
   SymbolicIOField "SIO_TL_BitNo" at 358,40 size 160x30; TextOff '0'; TextOn '1'; TextList "TL_BitNo"
      ProcessValue <- "D_Bits"
   TextField "Label_SIO_TL_BitNo" at 358,72 size 126x22; Text 'SIO_TL_BitNo'
   SymbolicIOField "SIO_TL_Value_Out" at 534,40 size 160x30; TextOff '0'; TextOn '1'; TextList "TL_Value"
      ProcessValue <- "D_TL"
   TextField "Label_SIO_TL_Value_Out" at 534,72 size 167x22; Text 'SIO_TL_Value_Out'
   GraphicIOField "GIO_GL_Value" at 710,40 size 120x80; PictureList "GL_Value"
      ProcessValue <- "D_TL"
   TextField "Label_GIO_GL_Value" at 710,122 size 129x22; Text 'GIO_GL_Value'
   GraphicIOField "GIO_GL_Bit" at 886,40 size 120x80; PictureList "GL_Bit"
      ProcessValue <- "D_Bool"
   TextField "Label_GIO_GL_Bit" at 886,122 size 106x22; Text 'GIO_GL_Bit'
   GraphicIOField "GIO_GL_BitNo" at 1062,40 size 120x80; PictureList "GL_BitNo"
      ProcessValue <- "D_Bits"
   TextField "Label_GIO_GL_BitNo" at 1062,122 size 129x22; Text 'GIO_GL_BitNo'
   GraphicIOField "GIO_GL_Value_Out" at 6,142 size 120x80; PictureList "GL_Value"
      ProcessValue <- "D_TL"
   TextField "Label_GIO_GL_Value_Out" at 6,224 size 170x22; Text 'GIO_GL_Value_Out'
   IOField "State" at 4,774 size 60x22; FormatPattern 9
      ProcessValue <- "D_State"
   Button "S1" at 70,774 size 40x22; TextOff 'S1'
      on Click: "SetS1"()
   Button "S2" at 114,774 size 40x22; TextOff 'S2'
      on Click: "SetS2"()
   Button "S3" at 158,774 size 40x22; TextOff 'S3'
      on Click: "SetS3"()
   Button "S4" at 202,774 size 40x22; TextOff 'S4'
      on Click: "SetS4"()
   Button "Next" at 1236,774 size 40x22; TextOff 'Next'
      on Click: ActivateScreen("C5_Buttons", 0)

Template "T_C05" 1280x800
   TextField "T_Title" at 8,6 size 185x21; Text 'Template T_C05 (header)'
   DateTimeField "T_Clock" at 1090,4 size 189x26

PopupScreen "Popup_C05" 300x200
   TextField "Pop_Title" at 10,10 size 224x22; Text 'Pop-up screen Popup_C05'
   GraphicView "Pop_Graphic" at 10,40 size 120x80; Picture "G_PNG"
   IOField "Pop_Value" at 150,60 size 120x30; FormatPattern s99999
      ProcessValue <- "D_Int"
   Button "Pop_Close" at 200,160 size 80x22; TextOff 'Close'
      on Click: function_efd93a16("Popup_C05", 200, 120, -1, -1, 1)

screen "C5_Structure" 1280x800, template "T_C05"
   Group "Group_A" at 10,50 size 300x87
   TextField "Label_Group_A (contains Group_B)" at 10,140 size 246x22; Text 'Group_A (contains Group_B)'
   TextField "Layer0_Text" at 352,52 size 69x22; Text 'Layer 0'
   TextField "Label_Layers 0-3 (layer 2 VisibleES false)" at 350,200 size 308x22; Text 'Layers 0-3 (layer 2 VisibleES false)'
   IOField "State" at 4,774 size 60x22; FormatPattern 9
      ProcessValue <- "D_State"
   Button "S1" at 70,774 size 40x22; TextOff 'S1'
      on Click: "SetS1"()
   Button "S2" at 114,774 size 40x22; TextOff 'S2'
      on Click: "SetS2"()
   Button "S3" at 158,774 size 40x22; TextOff 'S3'
      on Click: "SetS3"()
   Button "S4" at 202,774 size 40x22; TextOff 'S4'
      on Click: "SetS4"()
   Button "Popup" at 246,774 size 60x22; TextOff 'Popup'
      on Click: function_efd93a16("Popup_C05", 200, 120, -1, -1, 1)
   Button "SlideIn" at 310,774 size 60x22; TextOff 'Slide'
      on Click: "C5_ToggleSlideIn"()
   Button "Next" at 1236,774 size 40x22; TextOff 'Next'
      on Click: ActivateScreen("C5_GraphicView_1", 0)
   Group "Group_B" at 210,50 size 100x87
   TextField "GB_Text" at 210,115 size 77x22; Text 'Group_B'
   TextField "Layer1_Text" at 382,72 size 69x22; Text 'Layer 1'
   TextField "Layer2_Text" at 412,92 size 69x22; Text 'Layer 2'
   TextField "Layer3_Text" at 442,112 size 69x22; Text 'Layer 3'

screen "C6_Faceplates" 1280x800
   ScreenModuleView "FP_Dyn" at 10,10 size 300x150; ScreenModuleType ""; Guid_{11997190-83750} 'Tags D_Int D_Range D_Pct'
      Guid_{11997190-83886} <- "D_Int"
      Guid_{11997190-83896} <- "D_Range"
      Guid_{11997190-83898} <- "D_Pct"
      Guid_{11997190-83900} <- "D_Vis"
   TextField "Label_FP_Dyn" at 10,162 size 69x22; Text 'FP_Dyn'
   ScreenModuleView "FP_Static" at 330,10 size 300x150; ScreenModuleType ""; Guid_{11997190-83750} 'Static values'
   TextField "Label_FP_Static" at 330,162 size 87x22; Text 'FP_Static'
   ScreenModuleView "FP_Alt" at 10,186 size 300x150; ScreenModuleType ""; Guid_{11997190-83750} 'Tags D_SInt D_TL D_UInt'
      Guid_{11997190-83886} <- "D_SInt"
      Guid_{11997190-83896} <- "D_TL"
      Guid_{11997190-83898} <- "D_UInt"
      Guid_{11997190-83900} <- "D_En"
   TextField "Label_FP_Alt" at 10,338 size 61x22; Text 'FP_Alt'
   ScreenModuleView "FP_Move" at 330,186 size 300x150; ScreenModuleType ""; Guid_{11997190-83750} 'Moved by D_Pct'
      Guid_{11997190-83886} <- "D_Int"
      Guid_{11997190-83896} <- "D_Range"
      Guid_{11997190-83898} <- "D_Pct"
      Guid_{11997190-83900} <- "D_Vis"
      HorizontalMovement <- "D_Pct"
   TextField "Label_FP_Move" at 330,338 size 81x22; Text 'FP_Move'
   IOField "State" at 4,774 size 60x22; FormatPattern 9
      ProcessValue <- "D_State"
   Button "S1" at 70,774 size 40x22; TextOff 'S1'
      on Click: "SetS1"()
   Button "S2" at 114,774 size 40x22; TextOff 'S2'
      on Click: "SetS2"()
   Button "S3" at 158,774 size 40x22; TextOff 'S3'
      on Click: "SetS3"()
   Button "S4" at 202,774 size 40x22; TextOff 'S4'
      on Click: "SetS4"()
   Button "Next" at 1236,774 size 40x22; TextOff 'Next'
      on Click: ActivateScreen("C6_Faceplates", 0)

VB script "SetS1"
   SmartTags("D_State") = 1
   SmartTags("D_Bool") = False
   SmartTags("D_SInt") = -128
   SmartTags("D_Int") = -32768
   SmartTags("D_DInt") = -2147483648
   SmartTags("D_USInt") = 0
   SmartTags("D_UInt") = 0
   SmartTags("D_UDInt") = 0
   SmartTags("D_Real") = -999.999
   SmartTags("D_LReal") = -0.00000015
   SmartTags("D_String") = ""
   SmartTags("D_DateTime") = DateSerial(1990, 1, 1) + TimeSerial(0, 0, 0)
   SmartTags("D_Pct") = 0
   SmartTags("D_Range") = 5
   SmartTags("D_Bits") = 1
   SmartTags("D_Vis") = False
   SmartTags("D_En") = False
   SmartTags("D_X") = 10
   SmartTags("D_Y") = 10
   SmartTags("D_Max") = 100
   SmartTags("D_Min") = 0
   SmartTags("D_TL") = -5
   SmartTags("D_BarR") = -5

VB script "SetS2"
   SmartTags("D_State") = 2
   SmartTags("D_Bool") = True
   SmartTags("D_SInt") = 12
   SmartTags("D_Int") = 1234
   SmartTags("D_DInt") = 123456
   SmartTags("D_USInt") = 200
   SmartTags("D_UInt") = 40000
   SmartTags("D_UDInt") = 3000000000
   SmartTags("D_Real") = 3.14159
   SmartTags("D_LReal") = 2.718281828
   SmartTags("D_String") = "Hello World"
   SmartTags("D_DateTime") = DateSerial(2026, 11, 22) + TimeSerial(13, 45, 30)
   SmartTags("D_Pct") = 50
   SmartTags("D_Range") = 25
   SmartTags("D_Bits") = 2
   SmartTags("D_Vis") = True
   SmartTags("D_En") = True
   SmartTags("D_X") = 320
   SmartTags("D_Y") = 200
   SmartTags("D_Max") = 200
   SmartTags("D_Min") = -100
   SmartTags("D_TL") = 5
   SmartTags("D_BarR") = 0

VB script "SetS3"
   SmartTags("D_State") = 3
   SmartTags("D_Bool") = True
   SmartTags("D_SInt") = 127
   SmartTags("D_Int") = 32767
   SmartTags("D_DInt") = 2147483647
   SmartTags("D_USInt") = 255
   SmartTags("D_UInt") = 65535
   SmartTags("D_UDInt") = 4294967295
   SmartTags("D_Real") = 123456.789
   SmartTags("D_LReal") = 1E+300
   SmartTags("D_String") = "Ünïcödé äöüß ÄÖÜ € – long text that is wider than the field 0123456789 ABCDEFGHIJ"
   SmartTags("D_DateTime") = DateSerial(2099, 12, 31) + TimeSerial(23, 59, 59)
   SmartTags("D_Pct") = 100
   SmartTags("D_Range") = 75
   SmartTags("D_Bits") = 4
   SmartTags("D_Vis") = True
   SmartTags("D_En") = False
   SmartTags("D_X") = 853
   SmartTags("D_Y") = 400
   SmartTags("D_Max") = 50
   SmartTags("D_Min") = -50
   SmartTags("D_TL") = 10
   SmartTags("D_BarR") = 5

VB script "SetS4"
   SmartTags("D_State") = 4
   SmartTags("D_Bool") = False
   SmartTags("D_SInt") = -1
   SmartTags("D_Int") = -1
   SmartTags("D_DInt") = 0
   SmartTags("D_USInt") = 1
   SmartTags("D_UInt") = 1
   SmartTags("D_UDInt") = 1
   SmartTags("D_Real") = 0.0005
   SmartTags("D_LReal") = -0.0
   SmartTags("D_String") = "äöü ÄÖÜ ß"
   SmartTags("D_DateTime") = DateSerial(1970, 1, 1) + TimeSerial(0, 0, 0)
   SmartTags("D_Pct") = 150
   SmartTags("D_Range") = 200
   SmartTags("D_Bits") = 9
   SmartTags("D_Vis") = False
   SmartTags("D_En") = True
   SmartTags("D_X") = -20
   SmartTags("D_Y") = 0
   SmartTags("D_Max") = 100
   SmartTags("D_Min") = 0
   SmartTags("D_TL") = 50
   SmartTags("D_BarR") = 2.5

VB script "C5_ToggleSlideIn"
   cf6f4242-93bf-47b4-8281-e920249d00b8 GraphX_Slidein_Top, $3$hmiToggle$
*)

(* ===== HMI "HMI_RT_1" =====

ScreenModuleEditorView "FP-C05" 640x480
   Rectangle "FP_Status" at 20,20 size 60x40
      Appearance <- "FRange"
   IOField "FP_Value" at 100,20 size 100x30; FormatPattern s99999
      ProcessValue <- "FValue"
   Bar "FP_Bar" at 220,20 size 30x130; MinimumValue 0; MaximumValue 100
      ProcessValue <- "FPct"
   Circle "FP_Lamp" at 260,20 size 40x40
      Visibility <- "FVis"
   TextField "FP_Title" at 20,120 size 180x20; Text 'Faceplate FP_C05'
*)